Fanuc KAREL source: KT00681.KL

PROGRAM KT00681
%NOLOCKGROUP
VAR
  P1: JOINTPOS
  P2: JOINTPOS
  OUT: BOOLEAN
BEGIN
  OUT = NOT P1
END KT00681
